ABB RobotStudio station: q7n4-workcell.rspag

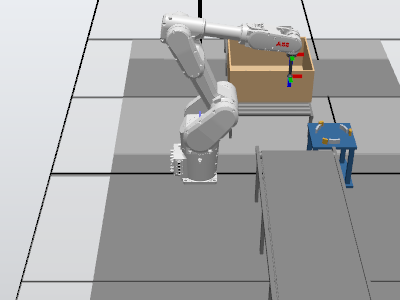
--- station ---
Station q7n4-initial-final015 (saved by RobotStudio 26.3.11794.0)
Controller System001
  mechanical unit ROB_1: IRB1300_7_140, 6 joints, base frame (0, 0, 0) mm
Layout (positions relative to the parent item):
  - IRB1300_7_140 [mechanism, from %ABB.RobotStudio.Models.IRB1300%\IRB1300_7_140__01.rslib] at (0, 0, 0) mm; joint values [0, -0.4958, 0.6435, 0, 1.4231, -3.1416] (rad or m)
  - InterimFixtureBase [part] at (850, 0, 0) mm, size 300 x 300 x 320 mm
  - PackingSupportRollers [part] at (500, 800, 0) mm, size 547.4 x 1396.2 x 49.2 mm
  - PackingSupportFrame [part] at (500, 800, 0) mm, size 587.9 x 1403 x 212.1 mm
  - InterimFixtureRadialGuides [part] at (850, 0, 350) mm, size 200.3 x 229.9 x 37 mm
  - InterimFixtureAnnularPads [part] at (850, 0, 350) mm, size 208.8 x 187.2 x 30 mm
  - SourcePart [part] at (600, -1730, 350) mm, size 226.4 x 215 x 150 mm
  - PackingCradle_PositiveY_BoxPart_1 [part] at (279.72, 680, 351.02) mm, rotated rx 0 ry 70 rz 0 deg, size 22.2 x 20.2 x 42 mm
  - PackingCradle_NegativeY_BoxPart_1 [part] at (279.72, 680, 351.02) mm, rotated rx 0 ry 70 rz 0 deg, size 22.2 x 20.2 x 42 mm
  - PackingCradle_PositiveY_BoxPart_2 [part] at (459.42, 680, 351.02) mm, rotated rx 0 ry 70 rz 0 deg, size 22.2 x 20.2 x 42 mm
  - PackingCradle_NegativeY_BoxPart_2 [part] at (459.42, 680, 351.02) mm, rotated rx 0 ry 70 rz 0 deg, size 22.2 x 20.2 x 42 mm
  - PackingCradle_PositiveY_BoxPart_3 [part] at (639.12, 680, 351.02) mm, rotated rx 0 ry 70 rz 0 deg, size 22.2 x 20.2 x 42 mm
  - PackingCradle_NegativeY_BoxPart_3 [part] at (639.12, 680, 351.02) mm, rotated rx 0 ry 70 rz 0 deg, size 22.2 x 20.2 x 42 mm
  - PackingCradle_PositiveY_BoxPart_4 [part] at (279.72, 920, 351.02) mm, rotated rx 0 ry 70 rz 0 deg, size 22.2 x 20.2 x 42 mm
  - PackingCradle_NegativeY_BoxPart_4 [part] at (279.72, 920, 351.02) mm, rotated rx 0 ry 70 rz 0 deg, size 22.2 x 20.2 x 42 mm
  - PackingCradle_PositiveY_BoxPart_5 [part] at (459.42, 920, 351.02) mm, rotated rx 0 ry 70 rz 0 deg, size 22.2 x 20.2 x 42 mm
  - PackingCradle_NegativeY_BoxPart_5 [part] at (459.42, 920, 351.02) mm, rotated rx 0 ry 70 rz 0 deg, size 22.2 x 20.2 x 42 mm
  - PackingCradle_PositiveY_BoxPart_6 [part] at (639.12, 920, 351.02) mm, rotated rx 0 ry 70 rz 0 deg, size 22.2 x 20.2 x 42 mm
  - PackingCradle_NegativeY_BoxPart_6 [part] at (639.12, 920, 351.02) mm, rotated rx 0 ry 70 rz 0 deg, size 22.2 x 20.2 x 42 mm
  - VacuumTool [part] at (550, 0, 900) mm, rotated rx 180 ry 0 rz 0 deg, size 60 x 60 x 150 mm
  - Floor [part] at (-600, -2100, -40) mm, size 2212.2 x 4114.7 x 59 mm
  - PackingBoxFloor [part] at (207.95, 537.5, 235) mm, size 584.1 x 525 x 15 mm
  - PackingBoxWall1 [part] at (207.95, 537.5, 250) mm, size 584.1 x 10 x 240 mm
  - PackingBoxWall2 [part] at (207.95, 1052.5, 250) mm, size 584.1 x 10 x 240 mm
  - PackingBoxWall3 [part] at (207.95, 547.5, 250) mm, size 10 x 505 x 240 mm
  - PackingBoxWall4 [part] at (782.05, 547.5, 250) mm, size 10 x 505 x 240 mm
  - ConveyorSurface [part] at (600, -500, 350) mm, size 445.5 x 1627.9 x 16.2 mm
  - ConveyorBeltReturn [part] at (600, -500, 350) mm, size 445.5 x 1627.9 x 16.2 mm
  - ConveyorBeltWraps [part] at (600, -500, 350) mm, size 443.7 x 1682.7 x 62.2 mm
  - ConveyorEndRollers [part] at (600, -500, 350) mm, size 472.1 x 1666.1 x 46.2 mm
  - ConveyorFrame [part] at (600, -500, 350) mm, size 501.9 x 1802.3 x 331.3 mm
Attachment: VacuumTool is attached to IRB1300_7_140 / Link6

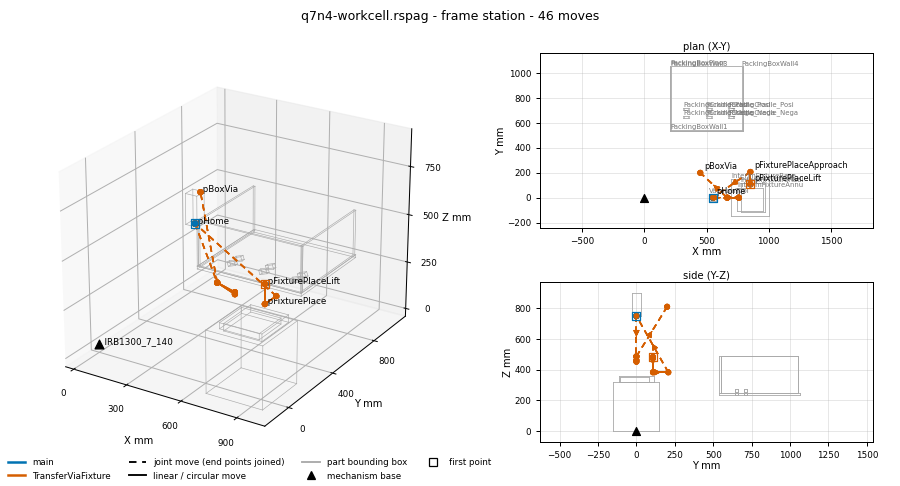
[picture p0: tool path of q7n4-workcell.rspag in frame station, 46 of 70 moves have a stored position in this frame; points joined in program order, loops and branches not executed]
--- Controller Data/System001/RAPID/TASK1/PROGMOD/MA6212_OnePiece014.modx ---
MODULE MA6212_OnePiece014
    ! One box of six actual parts; simulated camera data is read for each source.
    ! IRB1300 / OmniCore, TCP150. Fixture guides require vertical C2 lift.
    ! Camera offsets come from measured CAD pose, not the feed random-number table.
    ! First part is nominal; five following parts have independent random XY offsets.
    ! Actor capacity is six, with one empty-box acknowledgement before the batch.
    PERS bool single014ExecutionArmed:=FALSE;
    PERS num runId:=140301;
    PERS num cycleIndex:=1;
    PERS num slot:=0;
    PERS num dx:=0;
    PERS num dy:=0;
    PERS num stage:=0;
    PERS num runState:=0;
    PERS num completedCycles:=0;
    PERS num runAttempt:=0;
    PERS num lastError:=0;
    PERS num elapsed:=0;
    PERS bool motionSequenceComplete:=FALSE;
    PERS string runFile:="";
    PERS bool visionReady:=FALSE;
    PERS num visionSequence:=0;
    PERS num visionConsumedSequence:=0;
    PERS num visionDxMm:=0;
    PERS num visionDyMm:=0;
    PERS num visionVirtualTimeMs:=0;
    PERS string visionPartId:="";
    PERS string visionFrame:="";
    VAR num caseNumber;
    VAR robtarget measuredSourceContact;
    VAR robtarget measuredSourceLift;
    CONST speeddata vEmptyMoveJ:=[400,120,100,30];
    CONST speeddata vTravelCommission:=[400,120,100,30];
    CONST speeddata vApproachCommission:=[320,96,100,30];
    VAR clock cycleClock;
    VAR iodev cycleLog;
    VAR bool logOpen:=FALSE;
    VAR bool timingActive:=FALSE;
    PERS loaddata elbowLoadAtC1:=[2.5,[18.8352947,22.7884033,107.5],[0.706433772,-0.0308435638,-0.706433772,-0.0308435637],0.0135624012,0.0154981713,0.0231869125];
    PERS loaddata elbowLoadAtC2:=[2.5,[-18.8352947,1.30134567e-09,84.7115967],[0.521333805,0.477714416,-0.477714417,-0.521333805],0.0135624012,0.0154981713,0.0231869125];
    CONST robtarget sourceApproach:=[[602.9245075451499,-142.49999999999997,383.42727420088414],[0.5416752204197017,0.5416752204197021,-0.4545194776720435,0.4545194776720435],[0,-1,-1,0],[9E9,9E9,9E9,9E9,9E9,9E9]];
    CONST robtarget sourceContact:=[[602.9245075451499,-242.5,383.4272742008841],[0.5416752204197017,0.5416752204197021,-0.4545194776720435,0.4545194776720435],[-1,-2,-1,0],[9E9,9E9,9E9,9E9,9E9,9E9]];
    CONST robtarget sourceLift:=[[602.9245075451499,-242.5,483.4272742008841],[0.5416752204197017,0.5416752204197021,-0.4545194776720435,0.4545194776720435],[-1,-2,-1,0],[9E9,9E9,9E9,9E9,9E9,9E9]];
    CONST robtarget boxApproach:=[[345.55530043978405,680,810.1261272331978],[6.123233995736766E-17,1,1.232595164407831E-32,-3.015276387438861E-17],[0,0,-2,0],[9E9,9E9,9E9,9E9,9E9,9E9]];
    CONST robtarget boxContact:=[[345.55530043978405,680,470.12612723319785],[6.123233995736766E-17,1,1.232595164407831E-32,-3.015276387438861E-17],[0,0,-2,0],[9E9,9E9,9E9,9E9,9E9,9E9]];
    CONST robtarget pBoxApproachSix{6}:=[
        [[345.55530043978405,680,810.1261272331978],[6.123233995736766E-17,1,1.232595164407831E-32,-3.015276387438861E-17],[0,0,-2,0],[9E9,9E9,9E9,9E9,9E9,9E9]],
        [[525.2557954783952,680,810.1261272331978],[6.123233995736766E-17,1,1.232595164407831E-32,-3.015276387438861E-17],[0,0,-2,0],[9E9,9E9,9E9,9E9,9E9,9E9]],
        [[704.9562905170061,680,810.1261272331978],[6.123233995736766E-17,1,1.232595164407831E-32,-3.015276387438861E-17],[0,0,-2,0],[9E9,9E9,9E9,9E9,9E9,9E9]],
        [[345.55530043978405,920,810.1261272331978],[6.123233995736766E-17,1,1.232595164407831E-32,-3.015276387438861E-17],[0,0,-2,0],[9E9,9E9,9E9,9E9,9E9,9E9]],
        [[525.2557954783952,920,810.1261272331978],[6.123233995736766E-17,1,1.232595164407831E-32,-3.015276387438861E-17],[0,0,-2,0],[9E9,9E9,9E9,9E9,9E9,9E9]],
        [[704.9562905170061,920,810.1261272331978],[6.123233995736766E-17,1,1.232595164407831E-32,-3.015276387438861E-17],[0,0,-2,0],[9E9,9E9,9E9,9E9,9E9,9E9]]];
    CONST robtarget pBoxContactSix{6}:=[
        [[345.55530043978405,680,470.12612723319785],[6.123233995736766E-17,1,1.232595164407831E-32,-3.015276387438861E-17],[0,0,-2,0],[9E9,9E9,9E9,9E9,9E9,9E9]],
        [[525.2557954783952,680,470.12612723319785],[6.123233995736766E-17,1,1.232595164407831E-32,-3.015276387438861E-17],[0,0,-2,0],[9E9,9E9,9E9,9E9,9E9,9E9]],
        [[704.9562905170061,680,470.12612723319785],[6.123233995736766E-17,1,1.232595164407831E-32,-3.015276387438861E-17],[0,0,-2,0],[9E9,9E9,9E9,9E9,9E9,9E9]],
        [[345.55530043978405,920,470.12612723319785],[6.123233995736766E-17,1,1.232595164407831E-32,-3.015276387438861E-17],[0,0,-2,0],[9E9,9E9,9E9,9E9,9E9,9E9]],
        [[525.2557954783952,920,470.12612723319785],[6.123233995736766E-17,1,1.232595164407831E-32,-3.015276387438861E-17],[0,0,-2,0],[9E9,9E9,9E9,9E9,9E9,9E9]],
        [[704.9562905170061,920,470.12612723319785],[6.123233995736766E-17,1,1.232595164407831E-32,-3.015276387438861E-17],[0,0,-2,0],[9E9,9E9,9E9,9E9,9E9,9E9]]];
    CONST robtarget pHome:=[[550,0,750],[0,1,0,0],[0,0,-3,0],[9E9,9E9,9E9,9E9,9E9,9E9]];
    CONST robtarget pBoxVia:=[[450,200,810.1261272331978],[6.123233995736766E-17,1,1.232595164407831E-32,-3.015276387438861E-17],[0,0,-2,0],[9E9,9E9,9E9,9E9,9E9,9E9]];
    CONST robtarget pFixturePlaceLift:=[[852.9245075451499,107.5,483.4272742008841],[0.5416752204197017,0.5416752204197021,-0.4545194776720435,0.4545194776720435],[0,-1,-1,0],[9E9,9E9,9E9,9E9,9E9,9E9]];
    CONST robtarget pFixturePlace:=[[852.9245075451499,107.5,383.4272742008841],[0.5416752204197017,0.5416752204197021,-0.4545194776720435,0.4545194776720435],[0,-1,-1,0],[9E9,9E9,9E9,9E9,9E9,9E9]];
    CONST robtarget pFixturePlaceApproach:=[[852.9245075451499,207.50000000000003,383.42727420088414],[0.5416752204197017,0.5416752204197021,-0.4545194776720435,0.4545194776720435],[0,-1,-1,0],[9E9,9E9,9E9,9E9,9E9,9E9]];
    CONST robtarget pFixturePickApproach:=[[666.6229516856366,2.5411421082307575E-14,486.8080573302675],[5.015859645267624E-17,0.8191520442889917,-0,0.5735764363510463],[0,0,-3,1],[9E9,9E9,9E9,9E9,9E9,9E9]];
    CONST robtarget pFixturePick:=[[760.5922137642275,1.3164953090834047E-14,452.6060429977006],[5.015859645267624E-17,0.8191520442889917,-0,0.5735764363510463],[-1,0,-3,1],[9E9,9E9,9E9,9E9,9E9,9E9]];

    PROC main()
        IF NOT single014ExecutionArmed THEN
            TPWrite "OnePiece014 is not released for execution.";
            RETURN;
        ENDIF
        ! Consume one-shot permission before any possible motion.
        single014ExecutionArmed:=FALSE;
        IF runAttempt<>0 OR StrLen(runFile)=0 THEN
            TPWrite "Fresh module and unique HOME CSV runFile required.";
            Stop;
            RETURN;
        ENDIF
        runAttempt:=1;
        lastError:=0;
        completedCycles:=0;
        motionSequenceComplete:=FALSE;
        timingActive:=FALSE;
        elapsed:=0;
        stage:=0;
        runState:=1;
        Open "HOME:"+runFile,cycleLog\Append;
        logOpen:=TRUE;
        Write cycleLog,"run,cycle,dx_mm,dy_mm,slot,cycle_s,state,stage,err,"\NoNewLine;
        Write cycleLog,"vision_part_id,vision_seq,vision_virtual_ms";
        ConfJ \On;
        ConfL \On;
        SetDO doVacuum,0;
        WaitDI diVacuumOK,0\MaxTime:=2;
        SetDO doFeedRequest,0;
        WaitDI diFeedReady,0\MaxTime:=5;
        SetDO doBoxReset,0;
        WaitDI diBoxReady,0\MaxTime:=5;
        MoveJ pHome,vEmptyMoveJ,fine,tVacuum\WObj:=wobj0;
        ResetBox;
        FOR caseNumber FROM 1 TO 6 DO
            cycleIndex:=caseNumber;
            slot:=cycleIndex-1;
            visionReady:=FALSE;
            stage:=8;
            SetDO doFeedRequest,1;
            WaitDI diFeedReady,1\MaxTime:=5;
            WaitUntil visionReady AND visionSequence=cycleIndex\MaxTime:=5;
            IF visionSequence<=visionConsumedSequence OR visionFrame<>"station_world" OR
               StrLen(visionPartId)=0 OR Abs(visionDxMm)>5 OR Abs(visionDyMm)>5 THEN
                lastError:=-100;
                runState:=-1;
                WriteCycle "INVALID_VISION";
                Close cycleLog;
                logOpen:=FALSE;
                Stop;
                RETURN;
            ENDIF
            ! These measured offsets are the only source-position correction inputs.
            dx:=visionDxMm;
            dy:=visionDyMm;
            visionConsumedSequence:=visionSequence;
            visionReady:=FALSE;
            ClkReset cycleClock;
            ClkStart cycleClock;
            timingActive:=TRUE;
            TransferViaFixture;
            MoveJ pHome,vEmptyMoveJ,fine,tVacuum\WObj:=wobj0;
            ClkStop cycleClock;
            elapsed:=ClkRead(cycleClock);
            timingActive:=FALSE;
            WriteCycle "MOTION_SEQUENCE_RETURNED";
            SetDO doFeedRequest,0;
            WaitDI diFeedReady,0\MaxTime:=5;
            completedCycles:=cycleIndex;
        ENDFOR
        motionSequenceComplete:=TRUE;
        stage:=0;
        runState:=2;
        Close cycleLog;
        logOpen:=FALSE;
        Stop;
    ERROR
        lastError:=ERRNO;
        runState:=-1;
        motionSequenceComplete:=FALSE;
        IF timingActive THEN
            ClkStop cycleClock;
            elapsed:=ClkRead(cycleClock);
            timingActive:=FALSE;
        ENDIF
        IF logOpen THEN
            WriteCycle "ERROR";
            Close cycleLog;
            logOpen:=FALSE;
        ENDIF
        ! Preserve current vacuum/output state for inspection; no blind release/retry.
        RAISE;
    ENDPROC

    PROC TransferViaFixture()
        ! Current identity-wobj0/world layout: source branch uses measured Y.
        ! Root must still validate both branches with actual CalcJointT and paths.
        measuredSourceContact:=Offs(sourceContact,dx,dy,0);
        measuredSourceLift:=Offs(sourceLift,dx,dy,0);
        IF dy>0 THEN
            measuredSourceContact.robconf:=[0,-1,-1,0];
            measuredSourceLift.robconf:=[0,-1,-1,0];
        ELSE
            measuredSourceContact.robconf:=[-1,-2,-1,0];
            measuredSourceLift.robconf:=[-1,-2,-1,0];
        ENDIF
        stage:=10;
        MoveJ Offs(sourceApproach,dx,dy,0),vEmptyMoveJ,fine,tVacuum\WObj:=wobj0;
        MoveL measuredSourceContact,vApproachCommission,fine,tVacuum\WObj:=wobj0;
        WaitTime \InPos,0.25;
        SetDO doVacuum,1;
        WaitDI diVacuumOK,1\MaxTime:=2;
        GripLoad elbowLoadAtC1;
        MoveL measuredSourceLift,vApproachCommission,fine,tVacuum\WObj:=wobj0;
        stage:=20;
        MoveJ pFixturePlaceLift,vTravelCommission,fine,tVacuum\WObj:=wobj0;
        MoveL pFixturePlace,vApproachCommission,fine,tVacuum\WObj:=wobj0;
        WaitTime \InPos,0.25;
        SetDO doVacuum,0;
        WaitDI diVacuumOK,0\MaxTime:=2;
        GripLoad load0;
        MoveL pFixturePlaceApproach,vApproachCommission,fine,tVacuum\WObj:=wobj0;
        WaitTime 0.5;
        stage:=30;
        ! Empty-tool transit via existing Ready; actual MoveJ collision check still required.
        MoveJ pHome,vEmptyMoveJ,fine,tVacuum\WObj:=wobj0;
        MoveJ pFixturePickApproach,vEmptyMoveJ,fine,tVacuum\WObj:=wobj0;
        MoveL pFixturePick,vApproachCommission,fine,tVacuum\WObj:=wobj0;
        WaitTime \InPos,0.25;
        SetDO doVacuum,1;
        WaitDI diVacuumOK,1\MaxTime:=2;
        GripLoad elbowLoadAtC2;
        ! Offs is world+Z ONLY after Root verifies wobj0 axes equal station world.
        ! Clear the7mm guides by10mm, fine; next MoveL rises another24.202mm.
        MoveL Offs(pFixturePick,0,0,10),vApproachCommission,fine,tVacuum\WObj:=wobj0;
        MoveL pFixturePickApproach,vApproachCommission,fine,tVacuum\WObj:=wobj0;
        stage:=40;
        MoveJ pBoxVia,vTravelCommission,fine,tVacuum\WObj:=wobj0;
        MoveL pBoxApproachSix{slot+1},vApproachCommission,fine,tVacuum\WObj:=wobj0;
        MoveL pBoxContactSix{slot+1},vApproachCommission,fine,tVacuum\WObj:=wobj0;
        WaitTime \InPos,0.25;
        SetDO doVacuum,0;
        WaitDI diVacuumOK,0\MaxTime:=2;
        GripLoad load0;
        MoveL pBoxApproachSix{slot+1},vApproachCommission,fine,tVacuum\WObj:=wobj0;
        stage:=50;
    ENDPROC

    PROC ResetBox()
        stage:=5;
        SetDO doBoxReset,1;
        WaitDI diBoxReady,1\MaxTime:=5;
        SetDO doBoxReset,0;
        WaitDI diBoxReady,0\MaxTime:=5;
    ENDPROC

    PROC WriteCycle(string stateText)
        ! Each chunk stays within the RAPID string limit; together they form 12 CSV columns.
        Write cycleLog,NumToStr(runId,0)+","+NumToStr(cycleIndex,0)+","+NumToStr(dx,3)+","+
            NumToStr(dy,3)+","+NumToStr(slot,0)+","\NoNewLine;
        Write cycleLog,NumToStr(elapsed,4)+","+stateText+","+NumToStr(stage,0)+","+
            NumToStr(lastError,0)+","\NoNewLine;
        Write cycleLog,visionPartId+","\NoNewLine;
        Write cycleLog,NumToStr(visionConsumedSequence,0)+","+NumToStr(visionVirtualTimeMs,1);
    ENDPROC
ENDMODULE

--- Controller Data/System001/RAPID/TASK1/PROGMOD/MA6212_Tooling.modx ---
MODULE MA6212_Tooling
    PERS tooldata tVacuum:=[TRUE,[[0,0,150],[1,0,0,0]],[1,[0,0,75],[1,0,0,0],0.001,0.001,0.001]];
ENDMODULE

--- Controller Data/System001/HOME/basic6_281ccaa64d6f4af6b89ba81da6075728.mod ---
MODULE MA6212_OnePiece014
    ! One box of six actual parts; simulated camera data is read for each source.
    ! IRB1300 / OmniCore, TCP150. Fixture guides require vertical C2 lift.
    ! Camera offsets come from measured CAD pose, not the feed random-number table.
    ! First part is nominal; five following parts have independent random XY offsets.
    ! Actor capacity is six, with one empty-box acknowledgement before the batch.
    PERS bool single014ExecutionArmed:=FALSE;
    PERS num runId:=140301;
    PERS num cycleIndex:=1;
    PERS num slot:=0;
    PERS num dx:=0;
    PERS num dy:=0;
    PERS num stage:=0;
    PERS num runState:=0;
    PERS num completedCycles:=0;
    PERS num runAttempt:=0;
    PERS num lastError:=0;
    PERS num elapsed:=0;
    PERS bool motionSequenceComplete:=FALSE;
    PERS string runFile:="";
    PERS bool visionReady:=FALSE;
    PERS num visionSequence:=0;
    PERS num visionConsumedSequence:=0;
    PERS num visionDxMm:=0;
    PERS num visionDyMm:=0;
    PERS num visionVirtualTimeMs:=0;
    PERS string visionPartId:="";
    PERS string visionFrame:="";
    VAR num caseNumber;
    VAR robtarget measuredSourceContact;
    VAR robtarget measuredSourceLift;
    CONST speeddata vEmptyMoveJ:=[25,7.5,100,30];
    CONST speeddata vTravelCommission:=[25,7.5,100,30];
    CONST speeddata vApproachCommission:=[20,6,100,30];
    VAR clock cycleClock;
    VAR iodev cycleLog;
    VAR bool logOpen:=FALSE;
    VAR bool timingActive:=FALSE;
    PERS loaddata elbowLoadAtC1:=[2.5,[18.8352947,22.7884033,107.5],[0.706433772,-0.0308435638,-0.706433772,-0.0308435637],0.0135624012,0.0154981713,0.0231869125];
    PERS loaddata elbowLoadAtC2:=[2.5,[-18.8352947,1.30134567e-09,84.7115967],[0.521333805,0.477714416,-0.477714417,-0.521333805],0.0135624012,0.0154981713,0.0231869125];
    CONST robtarget sourceApproach:=[[602.9245075451499,-142.49999999999997,383.42727420088414],[0.5416752204197017,0.5416752204197021,-0.4545194776720435,0.4545194776720435],[0,-1,-1,0],[9E9,9E9,9E9,9E9,9E9,9E9]];
    CONST robtarget sourceContact:=[[602.9245075451499,-242.5,383.4272742008841],[0.5416752204197017,0.5416752204197021,-0.4545194776720435,0.4545194776720435],[-1,-2,-1,0],[9E9,9E9,9E9,9E9,9E9,9E9]];
    CONST robtarget sourceLift:=[[602.9245075451499,-242.5,483.4272742008841],[0.5416752204197017,0.5416752204197021,-0.4545194776720435,0.4545194776720435],[-1,-2,-1,0],[9E9,9E9,9E9,9E9,9E9,9E9]];
    CONST robtarget boxApproach:=[[345.55530043978405,680,810.1261272331978],[6.123233995736766E-17,1,1.232595164407831E-32,-3.015276387438861E-17],[0,0,-2,0],[9E9,9E9,9E9,9E9,9E9,9E9]];
    CONST robtarget boxContact:=[[345.55530043978405,680,470.12612723319785],[6.123233995736766E-17,1,1.232595164407831E-32,-3.015276387438861E-17],[0,0,-2,0],[9E9,9E9,9E9,9E9,9E9,9E9]];
    CONST robtarget pBoxApproachSix{6}:=[
        [[345.55530043978405,680,810.1261272331978],[6.123233995736766E-17,1,1.232595164407831E-32,-3.015276387438861E-17],[0,0,-2,0],[9E9,9E9,9E9,9E9,9E9,9E9]],
        [[525.2557954783952,680,810.1261272331978],[6.123233995736766E-17,1,1.232595164407831E-32,-3.015276387438861E-17],[0,0,-2,0],[9E9,9E9,9E9,9E9,9E9,9E9]],
        [[704.9562905170061,680,810.1261272331978],[6.123233995736766E-17,1,1.232595164407831E-32,-3.015276387438861E-17],[0,0,-2,0],[9E9,9E9,9E9,9E9,9E9,9E9]],
        [[345.55530043978405,920,810.1261272331978],[6.123233995736766E-17,1,1.232595164407831E-32,-3.015276387438861E-17],[0,0,-2,0],[9E9,9E9,9E9,9E9,9E9,9E9]],
        [[525.2557954783952,920,810.1261272331978],[6.123233995736766E-17,1,1.232595164407831E-32,-3.015276387438861E-17],[0,0,-2,0],[9E9,9E9,9E9,9E9,9E9,9E9]],
        [[704.9562905170061,920,810.1261272331978],[6.123233995736766E-17,1,1.232595164407831E-32,-3.015276387438861E-17],[0,0,-2,0],[9E9,9E9,9E9,9E9,9E9,9E9]]];
    CONST robtarget pBoxContactSix{6}:=[
        [[345.55530043978405,680,470.12612723319785],[6.123233995736766E-17,1,1.232595164407831E-32,-3.015276387438861E-17],[0,0,-2,0],[9E9,9E9,9E9,9E9,9E9,9E9]],
        [[525.2557954783952,680,470.12612723319785],[6.123233995736766E-17,1,1.232595164407831E-32,-3.015276387438861E-17],[0,0,-2,0],[9E9,9E9,9E9,9E9,9E9,9E9]],
        [[704.9562905170061,680,470.12612723319785],[6.123233995736766E-17,1,1.232595164407831E-32,-3.015276387438861E-17],[0,0,-2,0],[9E9,9E9,9E9,9E9,9E9,9E9]],
        [[345.55530043978405,920,470.12612723319785],[6.123233995736766E-17,1,1.232595164407831E-32,-3.015276387438861E-17],[0,0,-2,0],[9E9,9E9,9E9,9E9,9E9,9E9]],
        [[525.2557954783952,920,470.12612723319785],[6.123233995736766E-17,1,1.232595164407831E-32,-3.015276387438861E-17],[0,0,-2,0],[9E9,9E9,9E9,9E9,9E9,9E9]],
        [[704.9562905170061,920,470.12612723319785],[6.123233995736766E-17,1,1.232595164407831E-32,-3.015276387438861E-17],[0,0,-2,0],[9E9,9E9,9E9,9E9,9E9,9E9]]];
    CONST robtarget pHome:=[[550,0,750],[0,1,0,0],[0,0,-3,0],[9E9,9E9,9E9,9E9,9E9,9E9]];
    CONST robtarget pBoxVia:=[[450,200,810.1261272331978],[6.123233995736766E-17,1,1.232595164407831E-32,-3.015276387438861E-17],[0,0,-2,0],[9E9,9E9,9E9,9E9,9E9,9E9]];
    CONST robtarget pFixturePlaceLift:=[[852.9245075451499,107.5,483.4272742008841],[0.5416752204197017,0.5416752204197021,-0.4545194776720435,0.4545194776720435],[0,-1,-1,0],[9E9,9E9,9E9,9E9,9E9,9E9]];
    CONST robtarget pFixturePlace:=[[852.9245075451499,107.5,383.4272742008841],[0.5416752204197017,0.5416752204197021,-0.4545194776720435,0.4545194776720435],[0,-1,-1,0],[9E9,9E9,9E9,9E9,9E9,9E9]];
    CONST robtarget pFixturePlaceApproach:=[[852.9245075451499,207.50000000000003,383.42727420088414],[0.5416752204197017,0.5416752204197021,-0.4545194776720435,0.4545194776720435],[0,-1,-1,0],[9E9,9E9,9E9,9E9,9E9,9E9]];
    CONST robtarget pFixturePickApproach:=[[666.6229516856366,2.5411421082307575E-14,486.8080573302675],[5.015859645267624E-17,0.8191520442889917,-0,0.5735764363510463],[0,0,-3,1],[9E9,9E9,9E9,9E9,9E9,9E9]];
    CONST robtarget pFixturePick:=[[760.5922137642275,1.3164953090834047E-14,452.6060429977006],[5.015859645267624E-17,0.8191520442889917,-0,0.5735764363510463],[-1,0,-3,1],[9E9,9E9,9E9,9E9,9E9,9E9]];

    PROC main()
        IF NOT single014ExecutionArmed THEN
            TPWrite "OnePiece014 is not released for execution.";
            RETURN;
        ENDIF
        ! Consume one-shot permission before any possible motion.
        single014ExecutionArmed:=FALSE;
        IF runAttempt<>0 OR StrLen(runFile)=0 THEN
            TPWrite "Fresh module and unique HOME CSV runFile required.";
            Stop;
            RETURN;
        ENDIF
        runAttempt:=1;
        lastError:=0;
        completedCycles:=0;
        motionSequenceComplete:=FALSE;
        timingActive:=FALSE;
        elapsed:=0;
        stage:=0;
        runState:=1;
        Open "HOME:"+runFile,cycleLog\Append;
        logOpen:=TRUE;
        Write cycleLog,"run,cycle,dx_mm,dy_mm,slot,cycle_s,state,stage,err,"\NoNewLine;
        Write cycleLog,"vision_part_id,vision_seq,vision_virtual_ms";
        ConfJ \On;
        ConfL \On;
        SetDO doVacuum,0;
        WaitDI diVacuumOK,0\MaxTime:=2;
        SetDO doFeedRequest,0;
        WaitDI diFeedReady,0\MaxTime:=5;
        SetDO doBoxReset,0;
        WaitDI diBoxReady,0\MaxTime:=5;
        MoveJ pHome,vEmptyMoveJ,fine,tVacuum\WObj:=wobj0;
        ResetBox;
        FOR caseNumber FROM 1 TO 6 DO
            cycleIndex:=caseNumber;
            slot:=cycleIndex-1;
            visionReady:=FALSE;
            stage:=8;
            SetDO doFeedRequest,1;
            WaitDI diFeedReady,1\MaxTime:=5;
            WaitUntil visionReady AND visionSequence=cycleIndex\MaxTime:=5;
            IF visionSequence<=visionConsumedSequence OR visionFrame<>"station_world" OR
               StrLen(visionPartId)=0 OR Abs(visionDxMm)>5 OR Abs(visionDyMm)>5 THEN
                lastError:=-100;
                runState:=-1;
                WriteCycle "INVALID_VISION";
                Close cycleLog;
                logOpen:=FALSE;
                Stop;
                RETURN;
            ENDIF
            ! These measured offsets are the only source-position correction inputs.
            dx:=visionDxMm;
            dy:=visionDyMm;
            visionConsumedSequence:=visionSequence;
            visionReady:=FALSE;
            ClkReset cycleClock;
            ClkStart cycleClock;
            timingActive:=TRUE;
            TransferViaFixture;
            MoveJ pHome,vEmptyMoveJ,fine,tVacuum\WObj:=wobj0;
            ClkStop cycleClock;
            elapsed:=ClkRead(cycleClock);
            timingActive:=FALSE;
            WriteCycle "MOTION_SEQUENCE_RETURNED";
            SetDO doFeedRequest,0;
            WaitDI diFeedReady,0\MaxTime:=5;
            completedCycles:=cycleIndex;
        ENDFOR
        motionSequenceComplete:=TRUE;
        stage:=0;
        runState:=2;
        Close cycleLog;
        logOpen:=FALSE;
        Stop;
    ERROR
        lastError:=ERRNO;
        runState:=-1;
        motionSequenceComplete:=FALSE;
        IF timingActive THEN
            ClkStop cycleClock;
            elapsed:=ClkRead(cycleClock);
            timingActive:=FALSE;
        ENDIF
        IF logOpen THEN
            WriteCycle "ERROR";
            Close cycleLog;
            logOpen:=FALSE;
        ENDIF
        ! Preserve current vacuum/output state for inspection; no blind release/retry.
        RAISE;
    ENDPROC

    PROC TransferViaFixture()
        ! Current identity-wobj0/world layout: source branch uses measured Y.
        ! Root must still validate both branches with actual CalcJointT and paths.
        measuredSourceContact:=Offs(sourceContact,dx,dy,0);
        measuredSourceLift:=Offs(sourceLift,dx,dy,0);
        IF dy>0 THEN
            measuredSourceContact.robconf:=[0,-1,-1,0];
            measuredSourceLift.robconf:=[0,-1,-1,0];
        ELSE
            measuredSourceContact.robconf:=[-1,-2,-1,0];
            measuredSourceLift.robconf:=[-1,-2,-1,0];
        ENDIF
        stage:=10;
        MoveJ Offs(sourceApproach,dx,dy,0),vEmptyMoveJ,fine,tVacuum\WObj:=wobj0;
        MoveL measuredSourceContact,vApproachCommission,fine,tVacuum\WObj:=wobj0;
        WaitTime \InPos,0.25;
        SetDO doVacuum,1;
        WaitDI diVacuumOK,1\MaxTime:=2;
        GripLoad elbowLoadAtC1;
        MoveL measuredSourceLift,vApproachCommission,fine,tVacuum\WObj:=wobj0;
        stage:=20;
        MoveJ pFixturePlaceLift,vTravelCommission,fine,tVacuum\WObj:=wobj0;
        MoveL pFixturePlace,vApproachCommission,fine,tVacuum\WObj:=wobj0;
        WaitTime \InPos,0.25;
        SetDO doVacuum,0;
        WaitDI diVacuumOK,0\MaxTime:=2;
        GripLoad load0;
        MoveL pFixturePlaceApproach,vApproachCommission,fine,tVacuum\WObj:=wobj0;
        WaitTime 0.5;
        stage:=30;
        ! Empty-tool transit via existing Ready; actual MoveJ collision check still required.
        MoveJ pHome,vEmptyMoveJ,fine,tVacuum\WObj:=wobj0;
        MoveJ pFixturePickApproach,vEmptyMoveJ,fine,tVacuum\WObj:=wobj0;
        MoveL pFixturePick,vApproachCommission,fine,tVacuum\WObj:=wobj0;
        WaitTime \InPos,0.25;
        SetDO doVacuum,1;
        WaitDI diVacuumOK,1\MaxTime:=2;
        GripLoad elbowLoadAtC2;
        ! Offs is world+Z ONLY after Root verifies wobj0 axes equal station world.
        ! Clear the7mm guides by10mm, fine; next MoveL rises another24.202mm.
        MoveL Offs(pFixturePick,0,0,10),vApproachCommission,fine,tVacuum\WObj:=wobj0;
        MoveL pFixturePickApproach,vApproachCommission,fine,tVacuum\WObj:=wobj0;
        stage:=40;
        MoveJ pBoxVia,vTravelCommission,fine,tVacuum\WObj:=wobj0;
        MoveL pBoxApproachSix{slot+1},vApproachCommission,fine,tVacuum\WObj:=wobj0;
        MoveL pBoxContactSix{slot+1},vApproachCommission,fine,tVacuum\WObj:=wobj0;
        WaitTime \InPos,0.25;
        SetDO doVacuum,0;
        WaitDI diVacuumOK,0\MaxTime:=2;
        GripLoad load0;
        MoveL pBoxApproachSix{slot+1},vApproachCommission,fine,tVacuum\WObj:=wobj0;
        stage:=50;
    ENDPROC

    PROC ResetBox()
        stage:=5;
        SetDO doBoxReset,1;
        WaitDI diBoxReady,1\MaxTime:=5;
        SetDO doBoxReset,0;
        WaitDI diBoxReady,0\MaxTime:=5;
    ENDPROC

    PROC WriteCycle(string stateText)
        ! Each chunk stays within the RAPID string limit; together they form 12 CSV columns.
        Write cycleLog,NumToStr(runId,0)+","+NumToStr(cycleIndex,0)+","+NumToStr(dx,3)+","+
            NumToStr(dy,3)+","+NumToStr(slot,0)+","\NoNewLine;
        Write cycleLog,NumToStr(elapsed,4)+","+stateText+","+NumToStr(stage,0)+","+
            NumToStr(lastError,0)+","\NoNewLine;
        Write cycleLog,visionPartId+","\NoNewLine;
        Write cycleLog,NumToStr(visionConsumedSequence,0)+","+NumToStr(visionVirtualTimeMs,1);
    ENDPROC
ENDMODULE

--- Controller Data/System001/HOME/basic6_76193b5f05c9461c99fb0c85bbcaa0aa.mod ---
MODULE MA6212_OnePiece014
    ! One box of six actual parts; simulated camera data is read for each source.
    ! IRB1300 / OmniCore, TCP150. Fixture guides require vertical C2 lift.
    ! Camera offsets come from measured CAD pose, not the feed random-number table.
    ! First part is nominal; five following parts have independent random XY offsets.
    ! Actor capacity is six, with one empty-box acknowledgement before the batch.
    PERS bool single014ExecutionArmed:=FALSE;
    PERS num runId:=140301;
    PERS num cycleIndex:=1;
    PERS num slot:=0;
    PERS num dx:=0;
    PERS num dy:=0;
    PERS num stage:=0;
    PERS num runState:=0;
    PERS num completedCycles:=0;
    PERS num runAttempt:=0;
    PERS num lastError:=0;
    PERS num elapsed:=0;
    PERS bool motionSequenceComplete:=FALSE;
    PERS string runFile:="";
    PERS bool visionReady:=FALSE;
    PERS num visionSequence:=0;
    PERS num visionConsumedSequence:=0;
    PERS num visionDxMm:=0;
    PERS num visionDyMm:=0;
    PERS num visionVirtualTimeMs:=0;
    PERS string visionPartId:="";
    PERS string visionFrame:="";
    VAR num caseNumber;
    VAR robtarget measuredSourceContact;
    VAR robtarget measuredSourceLift;
    CONST speeddata vEmptyMoveJ:=[400,120,100,30];
    CONST speeddata vTravelCommission:=[400,120,100,30];
    CONST speeddata vApproachCommission:=[320,96,100,30];
    VAR clock cycleClock;
    VAR iodev cycleLog;
    VAR bool logOpen:=FALSE;
    VAR bool timingActive:=FALSE;
    PERS loaddata elbowLoadAtC1:=[2.5,[18.8352947,22.7884033,107.5],[0.706433772,-0.0308435638,-0.706433772,-0.0308435637],0.0135624012,0.0154981713,0.0231869125];
    PERS loaddata elbowLoadAtC2:=[2.5,[-18.8352947,1.30134567e-09,84.7115967],[0.521333805,0.477714416,-0.477714417,-0.521333805],0.0135624012,0.0154981713,0.0231869125];
    CONST robtarget sourceApproach:=[[602.9245075451499,-142.49999999999997,383.42727420088414],[0.5416752204197017,0.5416752204197021,-0.4545194776720435,0.4545194776720435],[0,-1,-1,0],[9E9,9E9,9E9,9E9,9E9,9E9]];
    CONST robtarget sourceContact:=[[602.9245075451499,-242.5,383.4272742008841],[0.5416752204197017,0.5416752204197021,-0.4545194776720435,0.4545194776720435],[-1,-2,-1,0],[9E9,9E9,9E9,9E9,9E9,9E9]];
    CONST robtarget sourceLift:=[[602.9245075451499,-242.5,483.4272742008841],[0.5416752204197017,0.5416752204197021,-0.4545194776720435,0.4545194776720435],[-1,-2,-1,0],[9E9,9E9,9E9,9E9,9E9,9E9]];
    CONST robtarget boxApproach:=[[345.55530043978405,680,810.1261272331978],[6.123233995736766E-17,1,1.232595164407831E-32,-3.015276387438861E-17],[0,0,-2,0],[9E9,9E9,9E9,9E9,9E9,9E9]];
    CONST robtarget boxContact:=[[345.55530043978405,680,470.12612723319785],[6.123233995736766E-17,1,1.232595164407831E-32,-3.015276387438861E-17],[0,0,-2,0],[9E9,9E9,9E9,9E9,9E9,9E9]];
    CONST robtarget pBoxApproachSix{6}:=[
        [[345.55530043978405,680,810.1261272331978],[6.123233995736766E-17,1,1.232595164407831E-32,-3.015276387438861E-17],[0,0,-2,0],[9E9,9E9,9E9,9E9,9E9,9E9]],
        [[525.2557954783952,680,810.1261272331978],[6.123233995736766E-17,1,1.232595164407831E-32,-3.015276387438861E-17],[0,0,-2,0],[9E9,9E9,9E9,9E9,9E9,9E9]],
        [[704.9562905170061,680,810.1261272331978],[6.123233995736766E-17,1,1.232595164407831E-32,-3.015276387438861E-17],[0,0,-2,0],[9E9,9E9,9E9,9E9,9E9,9E9]],
        [[345.55530043978405,920,810.1261272331978],[6.123233995736766E-17,1,1.232595164407831E-32,-3.015276387438861E-17],[0,0,-2,0],[9E9,9E9,9E9,9E9,9E9,9E9]],
        [[525.2557954783952,920,810.1261272331978],[6.123233995736766E-17,1,1.232595164407831E-32,-3.015276387438861E-17],[0,0,-2,0],[9E9,9E9,9E9,9E9,9E9,9E9]],
        [[704.9562905170061,920,810.1261272331978],[6.123233995736766E-17,1,1.232595164407831E-32,-3.015276387438861E-17],[0,0,-2,0],[9E9,9E9,9E9,9E9,9E9,9E9]]];
    CONST robtarget pBoxContactSix{6}:=[
        [[345.55530043978405,680,470.12612723319785],[6.123233995736766E-17,1,1.232595164407831E-32,-3.015276387438861E-17],[0,0,-2,0],[9E9,9E9,9E9,9E9,9E9,9E9]],
        [[525.2557954783952,680,470.12612723319785],[6.123233995736766E-17,1,1.232595164407831E-32,-3.015276387438861E-17],[0,0,-2,0],[9E9,9E9,9E9,9E9,9E9,9E9]],
        [[704.9562905170061,680,470.12612723319785],[6.123233995736766E-17,1,1.232595164407831E-32,-3.015276387438861E-17],[0,0,-2,0],[9E9,9E9,9E9,9E9,9E9,9E9]],
        [[345.55530043978405,920,470.12612723319785],[6.123233995736766E-17,1,1.232595164407831E-32,-3.015276387438861E-17],[0,0,-2,0],[9E9,9E9,9E9,9E9,9E9,9E9]],
        [[525.2557954783952,920,470.12612723319785],[6.123233995736766E-17,1,1.232595164407831E-32,-3.015276387438861E-17],[0,0,-2,0],[9E9,9E9,9E9,9E9,9E9,9E9]],
        [[704.9562905170061,920,470.12612723319785],[6.123233995736766E-17,1,1.232595164407831E-32,-3.015276387438861E-17],[0,0,-2,0],[9E9,9E9,9E9,9E9,9E9,9E9]]];
    CONST robtarget pHome:=[[550,0,750],[0,1,0,0],[0,0,-3,0],[9E9,9E9,9E9,9E9,9E9,9E9]];
    CONST robtarget pBoxVia:=[[450,200,810.1261272331978],[6.123233995736766E-17,1,1.232595164407831E-32,-3.015276387438861E-17],[0,0,-2,0],[9E9,9E9,9E9,9E9,9E9,9E9]];
    CONST robtarget pFixturePlaceLift:=[[852.9245075451499,107.5,483.4272742008841],[0.5416752204197017,0.5416752204197021,-0.4545194776720435,0.4545194776720435],[0,-1,-1,0],[9E9,9E9,9E9,9E9,9E9,9E9]];
    CONST robtarget pFixturePlace:=[[852.9245075451499,107.5,383.4272742008841],[0.5416752204197017,0.5416752204197021,-0.4545194776720435,0.4545194776720435],[0,-1,-1,0],[9E9,9E9,9E9,9E9,9E9,9E9]];
    CONST robtarget pFixturePlaceApproach:=[[852.9245075451499,207.50000000000003,383.42727420088414],[0.5416752204197017,0.5416752204197021,-0.4545194776720435,0.4545194776720435],[0,-1,-1,0],[9E9,9E9,9E9,9E9,9E9,9E9]];
    CONST robtarget pFixturePickApproach:=[[666.6229516856366,2.5411421082307575E-14,486.8080573302675],[5.015859645267624E-17,0.8191520442889917,-0,0.5735764363510463],[0,0,-3,1],[9E9,9E9,9E9,9E9,9E9,9E9]];
    CONST robtarget pFixturePick:=[[760.5922137642275,1.3164953090834047E-14,452.6060429977006],[5.015859645267624E-17,0.8191520442889917,-0,0.5735764363510463],[-1,0,-3,1],[9E9,9E9,9E9,9E9,9E9,9E9]];

    PROC main()
        IF NOT single014ExecutionArmed THEN
            TPWrite "OnePiece014 is not released for execution.";
            RETURN;
        ENDIF
        ! Consume one-shot permission before any possible motion.
        single014ExecutionArmed:=FALSE;
        IF runAttempt<>0 OR StrLen(runFile)=0 THEN
            TPWrite "Fresh module and unique HOME CSV runFile required.";
            Stop;
            RETURN;
        ENDIF
        runAttempt:=1;
        lastError:=0;
        completedCycles:=0;
        motionSequenceComplete:=FALSE;
        timingActive:=FALSE;
        elapsed:=0;
        stage:=0;
        runState:=1;
        Open "HOME:"+runFile,cycleLog\Append;
        logOpen:=TRUE;
        Write cycleLog,"run,cycle,dx_mm,dy_mm,slot,cycle_s,state,stage,err,"\NoNewLine;
        Write cycleLog,"vision_part_id,vision_seq,vision_virtual_ms";
        ConfJ \On;
        ConfL \On;
        SetDO doVacuum,0;
        WaitDI diVacuumOK,0\MaxTime:=2;
        SetDO doFeedRequest,0;
        WaitDI diFeedReady,0\MaxTime:=5;
        SetDO doBoxReset,0;
        WaitDI diBoxReady,0\MaxTime:=5;
        MoveJ pHome,vEmptyMoveJ,fine,tVacuum\WObj:=wobj0;
        ResetBox;
        FOR caseNumber FROM 1 TO 6 DO
            cycleIndex:=caseNumber;
            slot:=cycleIndex-1;
            visionReady:=FALSE;
            stage:=8;
            SetDO doFeedRequest,1;
            WaitDI diFeedReady,1\MaxTime:=5;
            WaitUntil visionReady AND visionSequence=cycleIndex\MaxTime:=5;
            IF visionSequence<=visionConsumedSequence OR visionFrame<>"station_world" OR
               StrLen(visionPartId)=0 OR Abs(visionDxMm)>5 OR Abs(visionDyMm)>5 THEN
                lastError:=-100;
                runState:=-1;
                WriteCycle "INVALID_VISION";
                Close cycleLog;
                logOpen:=FALSE;
                Stop;
                RETURN;
            ENDIF
            ! These measured offsets are the only source-position correction inputs.
            dx:=visionDxMm;
            dy:=visionDyMm;
            visionConsumedSequence:=visionSequence;
            visionReady:=FALSE;
            ClkReset cycleClock;
            ClkStart cycleClock;
            timingActive:=TRUE;
            TransferViaFixture;
            MoveJ pHome,vEmptyMoveJ,fine,tVacuum\WObj:=wobj0;
            ClkStop cycleClock;
            elapsed:=ClkRead(cycleClock);
            timingActive:=FALSE;
            WriteCycle "MOTION_SEQUENCE_RETURNED";
            SetDO doFeedRequest,0;
            WaitDI diFeedReady,0\MaxTime:=5;
            completedCycles:=cycleIndex;
        ENDFOR
        motionSequenceComplete:=TRUE;
        stage:=0;
        runState:=2;
        Close cycleLog;
        logOpen:=FALSE;
        Stop;
    ERROR
        lastError:=ERRNO;
        runState:=-1;
        motionSequenceComplete:=FALSE;
        IF timingActive THEN
            ClkStop cycleClock;
            elapsed:=ClkRead(cycleClock);
            timingActive:=FALSE;
        ENDIF
        IF logOpen THEN
            WriteCycle "ERROR";
            Close cycleLog;
            logOpen:=FALSE;
        ENDIF
        ! Preserve current vacuum/output state for inspection; no blind release/retry.
        RAISE;
    ENDPROC

    PROC TransferViaFixture()
        ! Current identity-wobj0/world layout: source branch uses measured Y.
        ! Root must still validate both branches with actual CalcJointT and paths.
        measuredSourceContact:=Offs(sourceContact,dx,dy,0);
        measuredSourceLift:=Offs(sourceLift,dx,dy,0);
        IF dy>0 THEN
            measuredSourceContact.robconf:=[0,-1,-1,0];
            measuredSourceLift.robconf:=[0,-1,-1,0];
        ELSE
            measuredSourceContact.robconf:=[-1,-2,-1,0];
            measuredSourceLift.robconf:=[-1,-2,-1,0];
        ENDIF
        stage:=10;
        MoveJ Offs(sourceApproach,dx,dy,0),vEmptyMoveJ,fine,tVacuum\WObj:=wobj0;
        MoveL measuredSourceContact,vApproachCommission,fine,tVacuum\WObj:=wobj0;
        WaitTime \InPos,0.25;
        SetDO doVacuum,1;
        WaitDI diVacuumOK,1\MaxTime:=2;
        GripLoad elbowLoadAtC1;
        MoveL measuredSourceLift,vApproachCommission,fine,tVacuum\WObj:=wobj0;
        stage:=20;
        MoveJ pFixturePlaceLift,vTravelCommission,fine,tVacuum\WObj:=wobj0;
        MoveL pFixturePlace,vApproachCommission,fine,tVacuum\WObj:=wobj0;
        WaitTime \InPos,0.25;
        SetDO doVacuum,0;
        WaitDI diVacuumOK,0\MaxTime:=2;
        GripLoad load0;
        MoveL pFixturePlaceApproach,vApproachCommission,fine,tVacuum\WObj:=wobj0;
        WaitTime 0.5;
        stage:=30;
        ! Empty-tool transit via existing Ready; actual MoveJ collision check still required.
        MoveJ pHome,vEmptyMoveJ,fine,tVacuum\WObj:=wobj0;
        MoveJ pFixturePickApproach,vEmptyMoveJ,fine,tVacuum\WObj:=wobj0;
        MoveL pFixturePick,vApproachCommission,fine,tVacuum\WObj:=wobj0;
        WaitTime \InPos,0.25;
        SetDO doVacuum,1;
        WaitDI diVacuumOK,1\MaxTime:=2;
        GripLoad elbowLoadAtC2;
        ! Offs is world+Z ONLY after Root verifies wobj0 axes equal station world.
        ! Clear the7mm guides by10mm, fine; next MoveL rises another24.202mm.
        MoveL Offs(pFixturePick,0,0,10),vApproachCommission,fine,tVacuum\WObj:=wobj0;
        MoveL pFixturePickApproach,vApproachCommission,fine,tVacuum\WObj:=wobj0;
        stage:=40;
        MoveJ pBoxVia,vTravelCommission,fine,tVacuum\WObj:=wobj0;
        MoveL pBoxApproachSix{slot+1},vApproachCommission,fine,tVacuum\WObj:=wobj0;
        MoveL pBoxContactSix{slot+1},vApproachCommission,fine,tVacuum\WObj:=wobj0;
        WaitTime \InPos,0.25;
        SetDO doVacuum,0;
        WaitDI diVacuumOK,0\MaxTime:=2;
        GripLoad load0;
        MoveL pBoxApproachSix{slot+1},vApproachCommission,fine,tVacuum\WObj:=wobj0;
        stage:=50;
    ENDPROC

    PROC ResetBox()
        stage:=5;
        SetDO doBoxReset,1;
        WaitDI diBoxReady,1\MaxTime:=5;
        SetDO doBoxReset,0;
        WaitDI diBoxReady,0\MaxTime:=5;
    ENDPROC

    PROC WriteCycle(string stateText)
        ! Each chunk stays within the RAPID string limit; together they form 12 CSV columns.
        Write cycleLog,NumToStr(runId,0)+","+NumToStr(cycleIndex,0)+","+NumToStr(dx,3)+","+
            NumToStr(dy,3)+","+NumToStr(slot,0)+","\NoNewLine;
        Write cycleLog,NumToStr(elapsed,4)+","+stateText+","+NumToStr(stage,0)+","+
            NumToStr(lastError,0)+","\NoNewLine;
        Write cycleLog,visionPartId+","\NoNewLine;
        Write cycleLog,NumToStr(visionConsumedSequence,0)+","+NumToStr(visionVirtualTimeMs,1);
    ENDPROC
ENDMODULE

--- Controller Data/System001/HOME/bootstrap014_6238bf105b8841babcbf657d91507fdb.mod ---
MODULE MA6212_Bootstrap014
    ! Candidate only; root must run the no-motion probe before the one MoveJ.
    CONST robtarget pReady014:=[[550,0,750],[0,1,0,0],[0,0,-3,0],[9E9,9E9,9E9,9E9,9E9,9E9]];
    CONST speeddata vBootstrap014:=[50,15,50,15];
    PERS bool motionArmed014:=FALSE;
    PERS bool probeCompleted014:=FALSE;
    PERS jointtarget readyJoints014:=[[0,0,0,0,0,0],[9E9,9E9,9E9,9E9,9E9,9E9]];
    PERS bool bootstrapAttempted014:=FALSE;
    PERS bool bootstrapCompleted014:=FALSE;
    PROC ProbeReady()
        readyJoints014:=CalcJointT(pReady014,tVacuum\WObj:=wobj0);
        probeCompleted014:=TRUE;
    ENDPROC
    PROC main()
        IF NOT motionArmed014 THEN
            ProbeReady;
            RETURN;
        ENDIF
        motionArmed014:=FALSE;
        IF NOT probeCompleted014 OR bootstrapAttempted014 THEN
            Stop;
            RETURN;
        ENDIF
        bootstrapAttempted014:=TRUE;
        ConfJ \On;
        GripLoad load0;
        MoveJ pReady014,vBootstrap014,fine,tVacuum\WObj:=wobj0;
        bootstrapCompleted014:=TRUE;
    ENDPROC
ENDMODULE

--- Controller Data/System001/HOME/bootstrap014_80a957812e4c435d8e72ee8011df24e6.mod ---
MODULE MA6212_Bootstrap014
    ! Candidate only; root must run the no-motion probe before the one MoveJ.
    CONST robtarget pReady014:=[[550,0,750],[0,1,0,0],[0,0,-3,0],[9E9,9E9,9E9,9E9,9E9,9E9]];
    ! Startup transfer: TCP25mm/s, orientation7.5deg/s.
    ! The former50/15 run686 stopped at the unchanged tracking guard; this run still requires actual verification.
    CONST speeddata vBootstrap014:=[25,7.5,50,15];
    PERS bool motionArmed014:=FALSE;
    PERS bool probeCompleted014:=FALSE;
    PERS jointtarget readyJoints014:=[[0,0,0,0,0,0],[9E9,9E9,9E9,9E9,9E9,9E9]];
    PERS bool bootstrapAttempted014:=FALSE;
    PERS bool bootstrapCompleted014:=FALSE;
    PROC ProbeReady()
        readyJoints014:=CalcJointT(pReady014,tVacuum\WObj:=wobj0);
        probeCompleted014:=TRUE;
    ENDPROC
    PROC main()
        IF NOT motionArmed014 THEN
            ProbeReady;
            RETURN;
        ENDIF
        motionArmed014:=FALSE;
        IF NOT probeCompleted014 OR bootstrapAttempted014 THEN
            Stop;
            RETURN;
        ENDIF
        bootstrapAttempted014:=TRUE;
        ConfJ \On;
        GripLoad load0;
        MoveJ pReady014,vBootstrap014,fine,tVacuum\WObj:=wobj0;
        bootstrapCompleted014:=TRUE;
    ENDPROC
ENDMODULE

--- Controller Data/System001/HOME/onepiece014_7d4820d1d5cd4c5498cd76560c1027ac.mod ---
MODULE MA6212_OnePiece014
    ! One box of six actual parts; simulated camera data is read for each source.
    ! IRB1300 / OmniCore, TCP150. Fixture guides require vertical C2 lift.
    ! Camera offsets come from measured CAD pose, not the feed random-number table.
    ! First part is nominal; five following parts have independent random XY offsets.
    ! Actor capacity is six, with one empty-box acknowledgement before the batch.
    PERS bool single014ExecutionArmed:=FALSE;
    PERS num runId:=140301;
    PERS num cycleIndex:=1;
    PERS num slot:=0;
    PERS num dx:=0;
    PERS num dy:=0;
    PERS num stage:=0;
    PERS num runState:=0;
    PERS num completedCycles:=0;
    PERS num runAttempt:=0;
    PERS num lastError:=0;
    PERS num elapsed:=0;
    PERS bool motionSequenceComplete:=FALSE;
    PERS string runFile:="";
    PERS bool visionReady:=FALSE;
    PERS num visionSequence:=0;
    PERS num visionConsumedSequence:=0;
    PERS num visionDxMm:=0;
    PERS num visionDyMm:=0;
    PERS num visionVirtualTimeMs:=0;
    PERS string visionPartId:="";
    PERS string visionFrame:="";
    VAR num caseNumber;
    VAR robtarget measuredSourceContact;
    VAR robtarget measuredSourceLift;
    CONST speeddata vEmptyMoveJ:=[25,7.5,100,30];
    CONST speeddata vTravelCommission:=[25,7.5,100,30];
    CONST speeddata vApproachCommission:=[20,6,100,30];
    VAR clock cycleClock;
    VAR iodev cycleLog;
    VAR bool logOpen:=FALSE;
    VAR bool timingActive:=FALSE;
    PERS loaddata elbowLoadAtC1:=[2.5,[18.8352947,22.7884033,107.5],[0.706433772,-0.0308435638,-0.706433772,-0.0308435637],0.0135624012,0.0154981713,0.0231869125];
    PERS loaddata elbowLoadAtC2:=[2.5,[-18.8352947,1.30134567e-09,84.7115967],[0.521333805,0.477714416,-0.477714417,-0.521333805],0.0135624012,0.0154981713,0.0231869125];
    CONST robtarget sourceApproach:=[[602.9245075451499,-142.49999999999997,383.42727420088414],[0.5416752204197017,0.5416752204197021,-0.4545194776720435,0.4545194776720435],[0,-1,-1,0],[9E9,9E9,9E9,9E9,9E9,9E9]];
    CONST robtarget sourceContact:=[[602.9245075451499,-242.5,383.4272742008841],[0.5416752204197017,0.5416752204197021,-0.4545194776720435,0.4545194776720435],[-1,-2,-1,0],[9E9,9E9,9E9,9E9,9E9,9E9]];
    CONST robtarget sourceLift:=[[602.9245075451499,-242.5,483.4272742008841],[0.5416752204197017,0.5416752204197021,-0.4545194776720435,0.4545194776720435],[-1,-2,-1,0],[9E9,9E9,9E9,9E9,9E9,9E9]];
    CONST robtarget boxApproach:=[[345.55530043978405,680,810.1261272331978],[6.123233995736766E-17,1,1.232595164407831E-32,-3.015276387438861E-17],[0,0,-2,0],[9E9,9E9,9E9,9E9,9E9,9E9]];
    CONST robtarget boxContact:=[[345.55530043978405,680,470.12612723319785],[6.123233995736766E-17,1,1.232595164407831E-32,-3.015276387438861E-17],[0,0,-2,0],[9E9,9E9,9E9,9E9,9E9,9E9]];
    CONST robtarget pBoxApproachSix{6}:=[
        [[345.55530043978405,680,810.1261272331978],[6.123233995736766E-17,1,1.232595164407831E-32,-3.015276387438861E-17],[0,0,-2,0],[9E9,9E9,9E9,9E9,9E9,9E9]],
        [[525.2557954783952,680,810.1261272331978],[6.123233995736766E-17,1,1.232595164407831E-32,-3.015276387438861E-17],[0,0,-2,0],[9E9,9E9,9E9,9E9,9E9,9E9]],
        [[704.9562905170061,680,810.1261272331978],[6.123233995736766E-17,1,1.232595164407831E-32,-3.015276387438861E-17],[0,0,-2,0],[9E9,9E9,9E9,9E9,9E9,9E9]],
        [[345.55530043978405,920,810.1261272331978],[6.123233995736766E-17,1,1.232595164407831E-32,-3.015276387438861E-17],[0,0,-2,0],[9E9,9E9,9E9,9E9,9E9,9E9]],
        [[525.2557954783952,920,810.1261272331978],[6.123233995736766E-17,1,1.232595164407831E-32,-3.015276387438861E-17],[0,0,-2,0],[9E9,9E9,9E9,9E9,9E9,9E9]],
        [[704.9562905170061,920,810.1261272331978],[6.123233995736766E-17,1,1.232595164407831E-32,-3.015276387438861E-17],[0,0,-2,0],[9E9,9E9,9E9,9E9,9E9,9E9]]];
    CONST robtarget pBoxContactSix{6}:=[
        [[345.55530043978405,680,470.12612723319785],[6.123233995736766E-17,1,1.232595164407831E-32,-3.015276387438861E-17],[0,0,-2,0],[9E9,9E9,9E9,9E9,9E9,9E9]],
        [[525.2557954783952,680,470.12612723319785],[6.123233995736766E-17,1,1.232595164407831E-32,-3.015276387438861E-17],[0,0,-2,0],[9E9,9E9,9E9,9E9,9E9,9E9]],
        [[704.9562905170061,680,470.12612723319785],[6.123233995736766E-17,1,1.232595164407831E-32,-3.015276387438861E-17],[0,0,-2,0],[9E9,9E9,9E9,9E9,9E9,9E9]],
        [[345.55530043978405,920,470.12612723319785],[6.123233995736766E-17,1,1.232595164407831E-32,-3.015276387438861E-17],[0,0,-2,0],[9E9,9E9,9E9,9E9,9E9,9E9]],
        [[525.2557954783952,920,470.12612723319785],[6.123233995736766E-17,1,1.232595164407831E-32,-3.015276387438861E-17],[0,0,-2,0],[9E9,9E9,9E9,9E9,9E9,9E9]],
        [[704.9562905170061,920,470.12612723319785],[6.123233995736766E-17,1,1.232595164407831E-32,-3.015276387438861E-17],[0,0,-2,0],[9E9,9E9,9E9,9E9,9E9,9E9]]];
    CONST robtarget pHome:=[[550,0,750],[0,1,0,0],[0,0,-3,0],[9E9,9E9,9E9,9E9,9E9,9E9]];
    CONST robtarget pBoxVia:=[[450,200,810.1261272331978],[6.123233995736766E-17,1,1.232595164407831E-32,-3.015276387438861E-17],[0,0,-2,0],[9E9,9E9,9E9,9E9,9E9,9E9]];
    CONST robtarget pFixturePlaceLift:=[[852.9245075451499,107.5,483.4272742008841],[0.5416752204197017,0.5416752204197021,-0.4545194776720435,0.4545194776720435],[0,-1,-1,0],[9E9,9E9,9E9,9E9,9E9,9E9]];
    CONST robtarget pFixturePlace:=[[852.9245075451499,107.5,383.4272742008841],[0.5416752204197017,0.5416752204197021,-0.4545194776720435,0.4545194776720435],[0,-1,-1,0],[9E9,9E9,9E9,9E9,9E9,9E9]];
    CONST robtarget pFixturePlaceApproach:=[[852.9245075451499,207.50000000000003,383.42727420088414],[0.5416752204197017,0.5416752204197021,-0.4545194776720435,0.4545194776720435],[0,-1,-1,0],[9E9,9E9,9E9,9E9,9E9,9E9]];
    CONST robtarget pFixturePickApproach:=[[666.6229516856366,2.5411421082307575E-14,486.8080573302675],[5.015859645267624E-17,0.8191520442889917,-0,0.5735764363510463],[0,0,-3,1],[9E9,9E9,9E9,9E9,9E9,9E9]];
    CONST robtarget pFixturePick:=[[760.5922137642275,1.3164953090834047E-14,452.6060429977006],[5.015859645267624E-17,0.8191520442889917,-0,0.5735764363510463],[-1,0,-3,1],[9E9,9E9,9E9,9E9,9E9,9E9]];

    PROC main()
        IF NOT single014ExecutionArmed THEN
            TPWrite "OnePiece014 is not released for execution.";
            RETURN;
        ENDIF
        ! Consume one-shot permission before any possible motion.
        single014ExecutionArmed:=FALSE;
        IF runAttempt<>0 OR StrLen(runFile)=0 THEN
            TPWrite "Fresh module and unique HOME CSV runFile required.";
            Stop;
            RETURN;
        ENDIF
        runAttempt:=1;
        lastError:=0;
        completedCycles:=0;
        motionSequenceComplete:=FALSE;
        timingActive:=FALSE;
        elapsed:=0;
        stage:=0;
        runState:=1;
        Open "HOME:"+runFile,cycleLog\Append;
        logOpen:=TRUE;
        Write cycleLog,"run,cycle,dx_mm,dy_mm,slot,cycle_s,state,stage,err,vision_part_id,vision_seq,vision_virtual_ms";
        ConfJ \On;
        ConfL \On;
        SetDO doVacuum,0;
        WaitDI diVacuumOK,0\MaxTime:=2;
        SetDO doFeedRequest,0;
        WaitDI diFeedReady,0\MaxTime:=5;
        SetDO doBoxReset,0;
        WaitDI diBoxReady,0\MaxTime:=5;
        MoveJ pHome,vEmptyMoveJ,fine,tVacuum\WObj:=wobj0;
        ResetBox;
        FOR caseNumber FROM 1 TO 6 DO
            cycleIndex:=caseNumber;
            slot:=cycleIndex-1;
            visionReady:=FALSE;
            stage:=8;
            SetDO doFeedRequest,1;
            WaitDI diFeedReady,1\MaxTime:=5;
            WaitUntil visionReady AND visionSequence=cycleIndex\MaxTime:=5;
            IF visionSequence<=visionConsumedSequence OR visionFrame<>"station_world" OR
               StrLen(visionPartId)=0 OR Abs(visionDxMm)>5 OR Abs(visionDyMm)>5 THEN
                lastError:=-100;
                runState:=-1;
                WriteCycle "INVALID_VISION";
                Close cycleLog;
                logOpen:=FALSE;
                Stop;
                RETURN;
            ENDIF
            ! These measured offsets are the only source-position correction inputs.
            dx:=visionDxMm;
            dy:=visionDyMm;
            visionConsumedSequence:=visionSequence;
            visionReady:=FALSE;
            ClkReset cycleClock;
            ClkStart cycleClock;
            timingActive:=TRUE;
            TransferViaFixture;
            MoveJ pHome,vEmptyMoveJ,fine,tVacuum\WObj:=wobj0;
            ClkStop cycleClock;
            elapsed:=ClkRead(cycleClock);
            timingActive:=FALSE;
            WriteCycle "MOTION_SEQUENCE_RETURNED";
            SetDO doFeedRequest,0;
            WaitDI diFeedReady,0\MaxTime:=5;
            completedCycles:=cycleIndex;
        ENDFOR
        motionSequenceComplete:=TRUE;
        stage:=0;
        runState:=2;
        Close cycleLog;
        logOpen:=FALSE;
        Stop;
    ERROR
        lastError:=ERRNO;
        runState:=-1;
        motionSequenceComplete:=FALSE;
        IF timingActive THEN
            ClkStop cycleClock;
            elapsed:=ClkRead(cycleClock);
            timingActive:=FALSE;
        ENDIF
        IF logOpen THEN
            WriteCycle "ERROR";
            Close cycleLog;
            logOpen:=FALSE;
        ENDIF
        ! Preserve current vacuum/output state for inspection; no blind release/retry.
        RAISE;
    ENDPROC

    PROC TransferViaFixture()
        ! Current identity-wobj0/world layout: source branch uses measured Y.
        ! Root must still validate both branches with actual CalcJointT and paths.
        measuredSourceContact:=Offs(sourceContact,dx,dy,0);
        measuredSourceLift:=Offs(sourceLift,dx,dy,0);
        IF dy>0 THEN
            measuredSourceContact.robconf:=[0,-1,-1,0];
            measuredSourceLift.robconf:=[0,-1,-1,0];
        ELSE
            measuredSourceContact.robconf:=[-1,-2,-1,0];
            measuredSourceLift.robconf:=[-1,-2,-1,0];
        ENDIF
        stage:=10;
        MoveJ Offs(sourceApproach,dx,dy,0),vEmptyMoveJ,fine,tVacuum\WObj:=wobj0;
        MoveL measuredSourceContact,vApproachCommission,fine,tVacuum\WObj:=wobj0;
        WaitTime \InPos,0.25;
        SetDO doVacuum,1;
        WaitDI diVacuumOK,1\MaxTime:=2;
        GripLoad elbowLoadAtC1;
        MoveL measuredSourceLift,vApproachCommission,fine,tVacuum\WObj:=wobj0;
        stage:=20;
        MoveJ pFixturePlaceLift,vTravelCommission,fine,tVacuum\WObj:=wobj0;
        MoveL pFixturePlace,vApproachCommission,fine,tVacuum\WObj:=wobj0;
        WaitTime \InPos,0.25;
        SetDO doVacuum,0;
        WaitDI diVacuumOK,0\MaxTime:=2;
        GripLoad load0;
        MoveL pFixturePlaceApproach,vApproachCommission,fine,tVacuum\WObj:=wobj0;
        WaitTime 0.5;
        stage:=30;
        ! Empty-tool transit via existing Ready; actual MoveJ collision check still required.
        MoveJ pHome,vEmptyMoveJ,fine,tVacuum\WObj:=wobj0;
        MoveJ pFixturePickApproach,vEmptyMoveJ,fine,tVacuum\WObj:=wobj0;
        MoveL pFixturePick,vApproachCommission,fine,tVacuum\WObj:=wobj0;
        WaitTime \InPos,0.25;
        SetDO doVacuum,1;
        WaitDI diVacuumOK,1\MaxTime:=2;
        GripLoad elbowLoadAtC2;
        ! Offs is world+Z ONLY after Root verifies wobj0 axes equal station world.
        ! Clear the7mm guides by10mm, fine; next MoveL rises another24.202mm.
        MoveL Offs(pFixturePick,0,0,10),vApproachCommission,fine,tVacuum\WObj:=wobj0;
        MoveL pFixturePickApproach,vApproachCommission,fine,tVacuum\WObj:=wobj0;
        stage:=40;
        MoveJ pBoxVia,vTravelCommission,fine,tVacuum\WObj:=wobj0;
        MoveL pBoxApproachSix{slot+1},vApproachCommission,fine,tVacuum\WObj:=wobj0;
        MoveL pBoxContactSix{slot+1},vApproachCommission,fine,tVacuum\WObj:=wobj0;
        WaitTime \InPos,0.25;
        SetDO doVacuum,0;
        WaitDI diVacuumOK,0\MaxTime:=2;
        GripLoad load0;
        MoveL pBoxApproachSix{slot+1},vApproachCommission,fine,tVacuum\WObj:=wobj0;
        stage:=50;
    ENDPROC

    PROC ResetBox()
        stage:=5;
        SetDO doBoxReset,1;
        WaitDI diBoxReady,1\MaxTime:=5;
        SetDO doBoxReset,0;
        WaitDI diBoxReady,0\MaxTime:=5;
    ENDPROC

    PROC WriteCycle(string stateText)
        Write cycleLog,NumToStr(runId,0)+","+NumToStr(cycleIndex,0)+","+NumToStr(dx,3)+","+
            NumToStr(dy,3)+","+NumToStr(slot,0)+","+NumToStr(elapsed,4)+","+
            stateText+","+NumToStr(stage,0)+","+NumToStr(lastError,0)+","+
            visionPartId+","+NumToStr(visionConsumedSequence,0)+","+NumToStr(visionVirtualTimeMs,1);
    ENDPROC
ENDMODULE

--- Controller Data/System001/HOME/targetprobe014_1cfdf8ed2334466e879ebe563a134cbd.mod ---
MODULE MA6212_TargetProbe014
    ! Unarmed, single-attempt target calculation only; no motion or IO operations.
    ! Exact target definitions from the reviewed OnePiece014 source are retained.
    PERS bool probeArmed014:=FALSE;
    PERS bool probeAttempted014:=FALSE;
    PERS bool probeCompleted014:=FALSE;
    PERS num probeTargetIndex014:=0;
    PERS num probeError014:=0;
    CONST robtarget sourceApproach:=[[602.9245075451499,-142.49999999999997,383.42727420088414],[0.5416752204197017,0.5416752204197021,-0.4545194776720435,0.4545194776720435],[0,-1,-1,0],[9E9,9E9,9E9,9E9,9E9,9E9]];
    CONST robtarget sourceContact:=[[602.9245075451499,-242.5,383.4272742008841],[0.5416752204197017,0.5416752204197021,-0.4545194776720435,0.4545194776720435],[-1,-2,-1,0],[9E9,9E9,9E9,9E9,9E9,9E9]];
    CONST robtarget sourceLift:=[[602.9245075451499,-242.5,483.4272742008841],[0.5416752204197017,0.5416752204197021,-0.4545194776720435,0.4545194776720435],[-1,-2,-1,0],[9E9,9E9,9E9,9E9,9E9,9E9]];
    CONST robtarget boxApproach:=[[345.55530043978405,680,810.1261272331978],[6.123233995736766E-17,1,1.232595164407831E-32,-3.015276387438861E-17],[0,0,-2,0],[9E9,9E9,9E9,9E9,9E9,9E9]];
    CONST robtarget boxContact:=[[345.55530043978405,680,470.12612723319785],[6.123233995736766E-17,1,1.232595164407831E-32,-3.015276387438861E-17],[0,0,-2,0],[9E9,9E9,9E9,9E9,9E9,9E9]];
    CONST robtarget pHome:=[[550,0,750],[0,1,0,0],[0,0,-3,0],[9E9,9E9,9E9,9E9,9E9,9E9]];
    CONST robtarget pBoxVia:=[[450,200,810.1261272331978],[6.123233995736766E-17,1,1.232595164407831E-32,-3.015276387438861E-17],[0,0,-2,0],[9E9,9E9,9E9,9E9,9E9,9E9]];
    CONST robtarget pFixturePlaceLift:=[[852.9245075451499,107.5,483.4272742008841],[0.5416752204197017,0.5416752204197021,-0.4545194776720435,0.4545194776720435],[0,-1,-1,0],[9E9,9E9,9E9,9E9,9E9,9E9]];
    CONST robtarget pFixturePlace:=[[852.9245075451499,107.5,383.4272742008841],[0.5416752204197017,0.5416752204197021,-0.4545194776720435,0.4545194776720435],[0,-1,-1,0],[9E9,9E9,9E9,9E9,9E9,9E9]];
    CONST robtarget pFixturePlaceApproach:=[[852.9245075451499,207.50000000000003,383.42727420088414],[0.5416752204197017,0.5416752204197021,-0.4545194776720435,0.4545194776720435],[0,-1,-1,0],[9E9,9E9,9E9,9E9,9E9,9E9]];
    CONST robtarget pFixturePickApproach:=[[666.6229516856366,2.5411421082307575E-14,486.8080573302675],[5.015859645267624E-17,0.8191520442889917,-0,0.5735764363510463],[0,0,-3,1],[9E9,9E9,9E9,9E9,9E9,9E9]];
    CONST robtarget pFixturePick:=[[760.5922137642275,1.3164953090834047E-14,452.6060429977006],[5.015859645267624E-17,0.8191520442889917,-0,0.5735764363510463],[-1,0,-3,1],[9E9,9E9,9E9,9E9,9E9,9E9]];
    PERS jointtarget probeJoints01014:=[[0,0,0,0,0,0],[9E9,9E9,9E9,9E9,9E9,9E9]];
    PERS jointtarget probeJoints02014:=[[0,0,0,0,0,0],[9E9,9E9,9E9,9E9,9E9,9E9]];
    PERS jointtarget probeJoints03014:=[[0,0,0,0,0,0],[9E9,9E9,9E9,9E9,9E9,9E9]];
    PERS jointtarget probeJoints04014:=[[0,0,0,0,0,0],[9E9,9E9,9E9,9E9,9E9,9E9]];
    PERS jointtarget probeJoints05014:=[[0,0,0,0,0,0],[9E9,9E9,9E9,9E9,9E9,9E9]];
    PERS jointtarget probeJoints06014:=[[0,0,0,0,0,0],[9E9,9E9,9E9,9E9,9E9,9E9]];
    PERS jointtarget probeJoints07014:=[[0,0,0,0,0,0],[9E9,9E9,9E9,9E9,9E9,9E9]];
    PERS jointtarget probeJoints08014:=[[0,0,0,0,0,0],[9E9,9E9,9E9,9E9,9E9,9E9]];
    PERS jointtarget probeJoints09014:=[[0,0,0,0,0,0],[9E9,9E9,9E9,9E9,9E9,9E9]];
    PERS jointtarget probeJoints10014:=[[0,0,0,0,0,0],[9E9,9E9,9E9,9E9,9E9,9E9]];
    PERS jointtarget probeJoints11014:=[[0,0,0,0,0,0],[9E9,9E9,9E9,9E9,9E9,9E9]];
    PERS jointtarget probeJoints12014:=[[0,0,0,0,0,0],[9E9,9E9,9E9,9E9,9E9,9E9]];
    PERS jointtarget probeJoints13014:=[[0,0,0,0,0,0],[9E9,9E9,9E9,9E9,9E9,9E9]];

    PROC main()
        IF NOT probeArmed014 THEN
            RETURN;
        ENDIF
        probeArmed014:=FALSE;
        IF probeAttempted014 THEN
            RETURN;
        ENDIF
        probeAttempted014:=TRUE;
        probeTargetIndex014:=1;
        probeJoints01014:=CalcJointT(sourceApproach,tVacuum\WObj:=wobj0);
        probeTargetIndex014:=2;
        probeJoints02014:=CalcJointT(sourceContact,tVacuum\WObj:=wobj0);
        probeTargetIndex014:=3;
        probeJoints03014:=CalcJointT(sourceLift,tVacuum\WObj:=wobj0);
        probeTargetIndex014:=4;
        probeJoints04014:=CalcJointT(boxApproach,tVacuum\WObj:=wobj0);
        probeTargetIndex014:=5;
        probeJoints05014:=CalcJointT(boxContact,tVacuum\WObj:=wobj0);
        probeTargetIndex014:=6;
        probeJoints06014:=CalcJointT(pHome,tVacuum\WObj:=wobj0);
        probeTargetIndex014:=7;
        probeJoints07014:=CalcJointT(pBoxVia,tVacuum\WObj:=wobj0);
        probeTargetIndex014:=8;
        probeJoints08014:=CalcJointT(pFixturePlaceLift,tVacuum\WObj:=wobj0);
        probeTargetIndex014:=9;
        probeJoints09014:=CalcJointT(pFixturePlace,tVacuum\WObj:=wobj0);
        probeTargetIndex014:=10;
        probeJoints10014:=CalcJointT(pFixturePlaceApproach,tVacuum\WObj:=wobj0);
        probeTargetIndex014:=11;
        probeJoints11014:=CalcJointT(pFixturePickApproach,tVacuum\WObj:=wobj0);
        probeTargetIndex014:=12;
        probeJoints12014:=CalcJointT(pFixturePick,tVacuum\WObj:=wobj0);
        probeTargetIndex014:=13;
        probeJoints13014:=CalcJointT(Offs(pFixturePick,0,0,10),tVacuum\WObj:=wobj0);
        probeCompleted014:=TRUE;
        RETURN;
    ERROR
        probeError014:=ERRNO;
        RAISE;
    ENDPROC
ENDMODULE

--- Controller Data/System001/SYSPAR/EIO.cfg ---
EIO:CFG_1.0:7:0::
#
VIRTUAL_NETWORK:

      -Name "Virtual" -Label "Virtual Device Network"
#
EIO_SIGNAL:

      -Name "IIO_di1" -SignalType "DI" -Device "IntegratedIOInternalDevice"\
      -DeviceMap "0"

      -Name "IIO_di2" -SignalType "DI" -Device "IntegratedIOInternalDevice"\
      -DeviceMap "1"

      -Name "IIO_di3" -SignalType "DI" -Device "IntegratedIOInternalDevice"\
      -DeviceMap "2"

      -Name "IIO_di4" -SignalType "DI" -Device "IntegratedIOInternalDevice"\
      -DeviceMap "3"

      -Name "IIO_di5" -SignalType "DI" -Device "IntegratedIOInternalDevice"\
      -DeviceMap "4"

      -Name "IIO_di6" -SignalType "DI" -Device "IntegratedIOInternalDevice"\
      -DeviceMap "5"

      -Name "IIO_di7" -SignalType "DI" -Device "IntegratedIOInternalDevice"\
      -DeviceMap "6"

      -Name "IIO_di8" -SignalType "DI" -Device "IntegratedIOInternalDevice"\
      -DeviceMap "7"

      -Name "IIO_di9" -SignalType "DI" -Device "IntegratedIOInternalDevice"\
      -DeviceMap "8"

      -Name "IIO_di10" -SignalType "DI" -Device "IntegratedIOInternalDevice"\
      -DeviceMap "9"

      -Name "IIO_di11" -SignalType "DI" -Device "IntegratedIOInternalDevice"\
      -DeviceMap "10"

      -Name "IIO_di12" -SignalType "DI" -Device "IntegratedIOInternalDevice"\
      -DeviceMap "11"

      -Name "IIO_di13" -SignalType "DI" -Device "IntegratedIOInternalDevice"\
      -DeviceMap "12"

      -Name "IIO_di14" -SignalType "DI" -Device "IntegratedIOInternalDevice"\
      -DeviceMap "13"

      -Name "IIO_di15" -SignalType "DI" -Device "IntegratedIOInternalDevice"\
      -DeviceMap "14"

      -Name "IIO_di16" -SignalType "DI" -Device "IntegratedIOInternalDevice"\
      -DeviceMap "15"

      -Name "IIO_do1" -SignalType "DO" -Device "IntegratedIOInternalDevice"\
      -DeviceMap "0"

      -Name "IIO_do2" -SignalType "DO" -Device "IntegratedIOInternalDevice"\
      -DeviceMap "1"

      -Name "IIO_do3" -SignalType "DO" -Device "IntegratedIOInternalDevice"\
      -DeviceMap "2"

      -Name "IIO_do4" -SignalType "DO" -Device "IntegratedIOInternalDevice"\
      -DeviceMap "3"

      -Name "IIO_do5" -SignalType "DO" -Device "IntegratedIOInternalDevice"\
      -DeviceMap "4"

      -Name "IIO_do6" -SignalType "DO" -Device "IntegratedIOInternalDevice"\
      -DeviceMap "5"

      -Name "IIO_do7" -SignalType "DO" -Device "IntegratedIOInternalDevice"\
      -DeviceMap "6"

      -Name "IIO_do8" -SignalType "DO" -Device "IntegratedIOInternalDevice"\
      -DeviceMap "7"

      -Name "IIO_gi" -SignalType "GI" -Device "integratedIOInternalDevice"\
      -DeviceMap "0-15"

      -Name "IIO_go" -SignalType "GO" -Device "integratedIOInternalDevice"\
      -DeviceMap "0-7"

      -Name "doVacuum" -SignalType "DO" -Access "All"

      -Name "diVacuumOK" -SignalType "DI" -Access "All"

      -Name "doFeedRequest" -SignalType "DO" -Access "All"

      -Name "diFeedReady" -SignalType "DI" -Access "All"

      -Name "doBoxReset" -SignalType "DO" -Access "All"

      -Name "diBoxReady" -SignalType "DI" -Access "All"

#CTRL_SIGNATURE:KsnpBxAUe/tzJvfXWyI7e0+0cnNCoo+Sist6FhcOtHJc0TgCUhL25MmDNrwyhcym4G7/tTtcyouiwOkd2tb+ZA==

--- Controller Data/System001/SYSPAR/PROC.cfg ---
PROC:CFG_1.0:7:0::

#CTRL_SIGNATURE:ME6O1W5CcTNsBEKWlKE06Hmm8XTykqSSfFnrm2k/ZJntiigvytBOOaSy1bfU5RV5/dlBHVdEJQV2kY+8o/9uPw==
